(*
    Configuration of FB_PlcShutdown.
*)
TYPE ST_ShutdownCfg :
STRUCT
    DelayMs : REAL := 3000.0;   // at Cmd.Shutdown; ms, >= 0, rounded to whole seconds
END_STRUCT
END_TYPE

(* stored: Version 1.1.0.1
   DUT ST_ShutdownCfg: Id {53ef0def-3a59-4757-8d00-5a4f051f5979} *)
